(* PLC project Vn_op_bool_to_int, Beckhoff Automation GmbH TwinCAT PLC Control 3.5.13.21 *)
(* stored: creationDateTime 1970-01-01T00:00:00 *)

PROGRAM Vn_op_bool_to_int

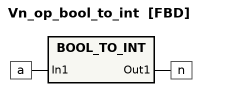
(* FBD diagram, written out as Structured Text *)
n := BOOL_TO_INT(a);
END_PROGRAM
